// TIA Portal V21 export
Screen "T09_IOMove"  1024x768, Number=29
  ScreenLayer 
    IOField "P_CraneX" at 0,0 size 100x30  DataFormat=Decimal, FormatPattern=s999999999.999, Mode=Output
      ProcessValue := Carried
      HorizontalMovementAnimation   RangeTo=9, Tag=CraneGX
